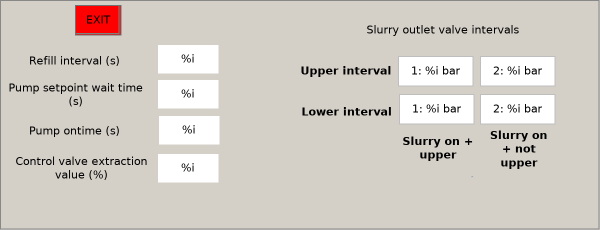
VISUALIZATION AutoExtractionParameterMenu  // 600x230
    Textfield (157,44 62x30), "%i", text variable: AutoExtractionParameterMenuBindings.refillIntervalTextField_TextVariable
        OnMouseDown: write the text variable via VisuDialogs.Numpad, min 1, max 999
    Label (23,39 103x44), "Refill interval (s)"
    Button (75,5 46x30), "EXIT", pressed state: NOT MainScreenBindings.autoExtractionParameterMenuButton_ToggleVariable
        toggle MainScreenBindings.autoExtractionParameterMenuButton_ToggleVariable
    Label (23,109 103x44), "Pump ontime (s)"
    Label (11,146 141x44), "Control valve extraction value (%)"
    Textfield (158,115 62x30), "%i", text variable: AutoExtractionParameterMenuBindings.pumpOnTimeTextField_TextVariable
        OnMouseDown: write the text variable via VisuDialogs.Numpad, min 1, max 5999
    Textfield (157,153 62x30), "%i", text variable: AutoExtractionParameterMenuBindings.controlValveOpeningValueTextField_TextVariable
        OnMouseDown: write the text variable via VisuDialogs.Numpad, min 1, max 5999
    Label (0,72 152x45), "Pump setpoint wait time (s)"
    Textfield (157,79 62x30), "%i", text variable: AutoExtractionParameterMenuBindings.pumpSetpointWaitTimeTextField_TextVariable
        OnMouseDown: write the text variable via VisuDialogs.Numpad, min 0, max 999
    Image (471,176 2x1), image: VisuSymbols.Symbols.ArrowBoldRight
    Label (296,49 100x44), "Upper interval"
    Label (297,90 100x44), "Lower interval"
    Textfield (398,56 75x30), "1: %i bar", text variable: MainScreenBindings.UpperIntervalSlurryOnUpperTextField_TextVariable
        OnMouseDown: write the text variable via VisuDialogs.Numpad, min -100, max 100
    Textfield (480,56 75x30), "2: %i bar", text variable: MainScreenBindings.UpperIntervalSlurryOnNotUpperTextField_TextVariable
        OnMouseDown: write the text variable via VisuDialogs.Numpad, min -100, max 100
    Textfield (399,94 75x30), "1: %i bar", text variable: MainScreenBindings.LowerIntervalSlurryOnUpperTextField_TextVariable
        OnMouseDown: write the text variable via VisuDialogs.Numpad, min -100, max 100
    Textfield (480,94 75x30), "2: %i bar", text variable: MainScreenBindings.LowerIntervalSlurryOnNotUpperTextField_TextVariable
        OnMouseDown: write the text variable via VisuDialogs.Numpad, min -100, max 100
    Label (399,126 78x44), "Slurry on + upper"
    Label (483,127 72x44), "Slurry on + not upper"
    Label (325,8 236x44), "Slurry outlet valve intervals"
END_VISUALIZATION

(* stored: Version 1.1.0.1, ProductVersion 3.1.4024.9
   Visu AutoExtractionParameterMenu: Id {88184fb8-5c74-471b-ba20-6c00e8dd02db} *)
